FUNCTION FC 1 : VOID
BEGIN
NETWORK
      A I 0.8
END_FUNCTION
